Staubli VAL3: io.pjx

--- io.pjx ---
Parameters version=s8.15.3Cs9_BS3337 stackSize=5000 millimeterUnit=true
Program file=getAnaIO.pgx
Program file=getDigIO.pgx
Program file=setAnaOutput.pgx
Program file=setDigOutput.pgx
Program file=start.pgx
Program file=stop.pgx
Program file=waitDigInput.pgx
Data file=io.dtx

--- io.dtx ---
mdesc mNomSpeed
public dio dInput[64]
public dio dOutput[64]
public aio aInput[16]
public aio aOutput[16]

--- start.pgx ---
program start()
begin
end

--- getAnaIO.pgx ---
public program getAnaIO(num x_nIndex, num& x_nValue, num& x_nResult)
  local string l_sDesc
  local string l_sPath
//读取模拟输入 aInput[x_nIndex]
//返回码 x_nResult: 0=正常  -1=索引越界  -2=该路未绑定物理通道(aioGet 会 runtime error，已提前拦截)
//注意：aInput 还没有 link（未做物理 IO 导入），此时读到的是恒 0 占位值，
//      必须先在 SRS 里完成物理 IO 导入，见 docs/05-IO绑定方法.md
begin
  x_nValue=0
  x_nResult=0

  //越界检查：合法下标 0..size(aInput)-1（手册 2.5.4，第31页 num size(*)）
  if (x_nIndex<0) or (x_nIndex>=size(aInput))
    x_nResult=-1
    return
  endIf

  //手册 3.6.1（第63页）：未 link 的 aio 参与运算会 runtime error，所以必须先 ioStatus
  //ioStatus(aio) 见手册 3.6.2（第64页），-1 = link 未定义
  if ioStatus(aInput[x_nIndex],l_sDesc,l_sPath)<0
    x_nResult=-2
    return
  endIf

  x_nValue=aioGet(aInput[x_nIndex])
end

--- getDigIO.pgx ---
public program getDigIO(num x_nIndex, bool& x_bValue, num& x_nResult)
  local string l_sDesc
  local string l_sPath
//读取数字输入 dInput[x_nIndex] 的电平
//返回码 x_nResult: 0=正常  -1=索引越界  -2=该位未绑定物理通道(ioStatus<0)
//注意：dInput 还没有 link（未做物理 IO 导入），此时读到的只是恒 0 占位值，
//      必须先在 SRS 里完成物理 IO 导入，见 docs/05-IO绑定方法.md
begin
  //先给默认值，任何提前 return 都不会把上一次的值留在引用参数里
  x_bValue=false
  x_nResult=0

  //越界检查：合法下标 0..size(dInput)-1（手册 2.5.4，第31页 num size(*)）
  if (x_nIndex<0) or (x_nIndex>=size(dInput))
    x_nResult=-1
    return
  endIf

  //未绑定物理通道时先拦截：手册 3.5.1（第59页）——未 link 的 dio 参与运算会触发 runtime error，
  //所以必须先 ioStatus 再读数；ioStatus 的 -1 含义见手册 3.5.3（第61页）：link 未定义
  if ioStatus(dInput[x_nIndex],l_sDesc,l_sPath)<0
    x_nResult=-2
    return
  endIf

  x_bValue=(dInput[x_nIndex]==true)
end

--- setAnaOutput.pgx ---
public program setAnaOutput(num x_nIndex, num x_nValue, num& x_nResult)
  local string l_sDesc
  local string l_sPath
//写模拟输出 aOutput[x_nIndex]
//返回码 x_nResult: 0=正常  -1=索引越界  -2=该路未绑定物理通道(aioSet 会 runtime error，已提前拦截)
//注意：aOutput 还没有 link（未做物理 IO 导入），此时写入不会作用到任何物理通道，
//      必须先在 SRS 里完成物理 IO 导入，见 docs/05-IO绑定方法.md
begin
  x_nResult=0

  //越界检查：合法下标 0..size(aOutput)-1（手册 2.5.4，第31页 num size(*)）
  if (x_nIndex<0) or (x_nIndex>=size(aOutput))
    x_nResult=-1
    return
  endIf

  //手册 3.6.1（第63页）：未 link 的 aio 参与运算会 runtime error，所以必须先 ioStatus
  if ioStatus(aOutput[x_nIndex],l_sDesc,l_sPath)<0
    x_nResult=-2
    return
  endIf

  aioSet(aOutput[x_nIndex],x_nValue)
end

--- setDigOutput.pgx ---
public program setDigOutput(num x_nIndex, bool x_bValue, num& x_nResult)
  local string l_sDesc
  local string l_sPath
//写数字输出 dOutput[x_nIndex]
//返回码 x_nResult: 0=正常  -1=索引越界  -2=该位未绑定物理通道(ioStatus<0，写入无效)
//注意：dOutput 还没有 link（未做物理 IO 导入），此时写入不会作用到任何物理点，
//      必须先在 SRS 里完成物理 IO 导入，见 docs/05-IO绑定方法.md
begin
  x_nResult=0

  //越界检查：合法下标 0..size(dOutput)-1（手册 2.5.4，第31页 num size(*)）
  if (x_nIndex<0) or (x_nIndex>=size(dOutput))
    x_nResult=-1
    return
  endIf

  //未绑定物理通道时先拦截：手册 3.5.2（第59页）——给未 link 的 dio 赋值会触发 runtime error
  if ioStatus(dOutput[x_nIndex],l_sDesc,l_sPath)<0
    x_nResult=-2
    return
  endIf

  dOutput[x_nIndex]=x_bValue
end

--- stop.pgx ---
program stop()
begin
end

--- waitDigInput.pgx ---
public program waitDigInput(num x_nIndex, bool x_bLevel, num x_nTimeout, bool& x_bDone, num& x_nResult)
  local string l_sDesc
  local string l_sPath
//等待数字输入 dInput[x_nIndex] 到达 x_bLevel 电平，带超时
//返回码 x_nResult: 0=已到达  -1=索引越界  -2=该位未绑定物理通道  -3=超时  -4=超时参数非法
//x_bDone=false 表示超时/未到达（唯一表示"等待失败"的语义位）
//注意：dInput 还没有 link（未做物理 IO 导入），此时读到的是恒 0，
//      等 true 一定等不到、只能超时；必须先在 SRS 里完成物理 IO 导入，见 docs/05-IO绑定方法.md
begin
  x_bDone=false
  x_nResult=0

  //越界检查：合法下标 0..size(dInput)-1（手册 2.5.4，第31页 num size(*)）
  if (x_nIndex<0) or (x_nIndex>=size(dInput))
    x_nResult=-1
    return
  endIf

  //未绑定物理通道时先拦截：手册 3.5.1（第59页）——未 link 的 dio 参与比较会触发 runtime error
  if ioStatus(dInput[x_nIndex],l_sDesc,l_sPath)<0
    x_nResult=-2
    return
  endIf

  //超时参数必须为正数，否则 watch() 会立刻返回 false，变成"假超时"
  if x_nTimeout<=0
    x_nResult=-4
    return
  endIf

  //watch() 手册 5 章（第103页）：条件在 nSeconds 内成立返回 true，超时返回 false。
  //相比 wait() 的好处是有超时，不会把任务永远挂住
  x_bDone=watch(dInput[x_nIndex]==x_bLevel,x_nTimeout)
  if x_bDone==false
    x_nResult=-3
  endIf
end
